(* IEC 61131-3 sources: ZPLC/conformance/com, 3 files *)

(* ---- com-002-a-failed-request-holds-error-while-en-stays-true.st ---- *)
PROGRAM Handshake
VAR
  Trigger AT %IX0.0 : BOOL;
  Link : MB_WRITE_COIL;
  Failed AT %QX0.0 : BOOL;
  Done AT %QX0.1 : BOOL;
  Busy AT %QX0.2 : BOOL;
  Code AT %QD1 : DINT;
END_VAR
  Link(EN := Trigger, PROTO := 1, SLAVE_ID := 1, ADDR := 0, COUNT := 1, VALUE := TRUE, HOST := '127.0.0.1', PORT := 502);
  Failed := Link.ERROR;
  Done := Link.DONE;
  Busy := Link.BUSY;
  Code := Link.STATUS;
END_PROGRAM

(* ---- com-002-a-request-is-one-for-each-rising-edge.st ---- *)
PROGRAM OneForEachEdge
VAR
  Trigger AT %IX0.0 : BOOL;
  Link : MQTT_PUBLISH;
  Edges AT %QW0 : INT;
  Previous : BOOL;
  Failed AT %QX2.0 : BOOL;
  Code AT %QD1 : DINT;
END_VAR
  Link(EN := Trigger, QOS := 0, RETAIN := FALSE, TOPIC := 'plant/a', PAYLOAD := 'x');
  Failed := Link.ERROR;
  Code := Link.STATUS;
  IF Link.ERROR AND NOT Previous THEN
    Edges := Edges + 1;
  END_IF;
  Previous := Link.ERROR;
END_PROGRAM

(* ---- com-005-string-arguments-of-a-block.st ---- *)
PROGRAM Strings
VAR
  Pub : MQTT_PUBLISH;
  Prov : AZURE_DPS_PROV;
  Rd : MB_READ_HREG;
  Name : STRING[20] := 'plant/line-7';
  TopicLen AT %QW0 : INT;
  PayloadLen AT %QW1 : INT;
  TopicOk AT %QX4.0 : BOOL;
  FromVariable AT %QW3 : INT;
  DeviceLen AT %QW4 : INT;
  HostLen AT %QW5 : INT;
  PortValue AT %QW6 : UINT;
END_VAR
  Pub(EN := FALSE, QOS := 1, RETAIN := FALSE, TOPIC := 'plant/a', PAYLOAD := 'hello');
  Prov(EN := FALSE, DEVICE_ID := Name);
  Rd(EN := FALSE, PROTO := 1, SLAVE_ID := 3, ADDR := 5, COUNT := 1, HOST := '10.0.0.5', PORT := 1502);
  TopicLen := LEN(Pub.TOPIC);
  PayloadLen := LEN(Pub.PAYLOAD);
  TopicOk := Pub.TOPIC = 'plant/a';
  FromVariable := LEN(Prov.DEVICE_ID);
  DeviceLen := LEN(Prov.ASSIGNED_HUB);
  HostLen := LEN(Rd.HOST);
  PortValue := Rd.PORT;
END_PROGRAM
